// TIA Portal V21 export
Screen "R04_BtnInv"  1024x768, Number=43, Template=Tpl
  ScreenLayer 
    Button "P_BtnInv" at 10,10 size 100x30  TextOff="BTN", TextOn="BTN"
      on Press: InvertBit(Tag := P_SwOn)
